SUBAPPLICATION MultipleOutputConnections
  (* Standard: 61499-1; Description: Copyright (c) 2026 Martin Erich Jobst This program and the accompanying materials are made available under the terms of the Eclipse Public License 2.0 which is available at https://www.eclipse.org/legal/epl-2.0/ SPDX-License-Identifier: EPL-2.0 *)
  (* Version 1.0, 2026-11-18, Martin Jobst *)
  PACKAGE lib::AdapterDeclaration;
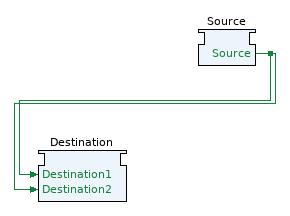
  SUBAPPLICATION Source
    PLUGS
      Source : lib::AdapterDeclaration::support::TestAdapter;
    END_PLUGS
  END_SUBAPPLICATION
  SUBAPPLICATION Destination
    SOCKETS
      Destination1 : lib::AdapterDeclaration::support::TestAdapter;
      Destination2 : lib::AdapterDeclaration::support::TestAdapter;
    END_SOCKETS
  END_SUBAPPLICATION
  ADAPTER_CONNECTIONS
    Source.Source TO Destination.Destination1;
    Source.Source TO Destination.Destination2;
  END_CONNECTIONS
END_SUBAPPLICATION
